// TIA Portal V20 export
Screen "Pop-up_PANEL_INITIALIZED_Popup"  800x400
  ScreenItem "Background" at 0,0 size 800x400  Type=HmiRectangle
  ScreenItem "Frame_Orange" at 3,3 size 794x394  Type=HmiRectangle
  ScreenItem "Button_Save" at 290,255 size 220x60  Type=HmiButton
  ScreenItem "Input_HMI_No" at 427,185 size 102x40  Type=HmiIOField
  ScreenItem "Text_Warning" at 200,85 size 400x70  Type=HmiTextBox
  ScreenItem "Text_HMI_No" at 272,185 size 150x40  Type=HmiTextBox
